// TIA Portal V20 export
// export: Created 2026-10-19T18:45:15.467375Z, ExportSetting None, DisplayName Totally Integrated Automation Portal, DisplayVersion V20 Update 6, DisplayName TIA Portal Openness, DisplayVersion V20 Update 6, DisplayName TIA Portal Version Control Interface, DisplayVersion V20 Update 6, DisplayName SINAMICS Startdrive Advanced, DisplayVersion V20 SP1, DisplayName SINAMICS Startdrive G130, G150, S120, S150, SINAMICS MV, G220, S200, S210, DisplayVersion V20 SP1, DisplayName SINAMICS Startdrive G110M, G120, G120C, G120D, G120P, G115D, DisplayVersion V20 SP1, DisplayName STEP 7 Professional, DisplayVersion V20 Update 6, DisplayName STEP 7 Safety, DisplayVersion V20 Update 2, DisplayName WinCC Basic/Comfort/Advanced, DisplayVersion V20 Update 6, DisplayName WinCC Unified, DisplayVersion V20 Update 6
VAR_GLOBAL   // PLC tag table "Screens"
   Main_OrderTable_Selected AT %MW114 : UInt;
   Settings_System_Selected AT %MW148 : UInt;
   Clear_OT AT %M154.0 : Bool;
   "Charger 1" AT %M154.1 : Bool;
   "Charger 2" AT %M154.2 : Bool;
   "Charger 3" AT %M154.3 : Bool;
   Shuttle_Level_Selected AT %MW112 : UInt;
   Charge_Shuttle_Commands AT %M136.0 : Bool;
   HMI_Box_Connected_4 AT %MW182 : Int;
   HMI_Box_Connected_5 AT %MW184 : Int;
   HMI_Box_Connected_3 AT %MW174 : Int;
   HMI_Box_Connected_2 AT %MW162 : Int;
   HMI_Box_Connected_1 AT %MW152 : Int;
   Shuttle_Level_EStop AT %M188.0 : Bool;
   Shuttle_EStop_All AT %M190.0 : Bool;
   All_In_Automatic_Buffers_2 AT %M510.5 : Bool;
   Automatic_Button_Buffers_1 AT %M510.6 : Bool;
   All_In_Automatic_Buffers_1 AT %M510.4 : Bool;
   Automatic_Button_Buffers_2 AT %M511.0 : Bool;
   Automatic_Button_VTD_2 AT %M510.7 : Bool;
   Automatic_Button_VTD_1 AT %M510.0 : Bool;
   All_In_Automatic_VTD_1 AT %M510.1 : Bool;
   All_In_Automatic_VTD_2 AT %M510.3 : Bool;
END_VAR
